TYPE "ST_ModuleTiming"
VERSION : 0.1
   STRUCT
      "LastCmdTime" : Time;
      "Rows" : Array[1..8] of "ST_TimingRow";
      "Truncated" : Bool;
   END_STRUCT;
END_TYPE
